(* IEC 61131-3 sources: PortalRobot/Portal_robot/Device/application/ST/ST_MULTI_TYPE, 4 files *)

(* ---- ST_MULTI_TYPE_COMMAND.st ---- *)
TYPE ST_MULTI_TYPE_COMMAND :
STRUCT
	{attribute 'symbol' := 'read'}
	xSetTypeCount         : BOOL; // Импульс изменения количества типов
	uiRequestedTypeCount : UINT; // Требуемое количество типов, 1..3
	{attribute 'symbol' := 'read'}
	xSetMachineType       : BOOL; // Импульс назначения типа станку
	uiRequestedMachine   : UINT; // Номер редактируемого станка, 1..3
	uiRequestedMachineType : UINT; // Тип, назначаемый станку
	{attribute 'symbol' := 'read'}
	xSetSlotType          : BOOL; // Импульс назначения типа слоту
	uiRequestedSlot      : UINT; // Номер редактируемого слота
	uiRequestedSlotType  : UINT; // Тип, назначаемый слоту
	{attribute 'symbol' := 'read'}
	xAutoDistribute      : BOOL; // Импульс распределения слотов пропорционально станкам
END_STRUCT
END_TYPE

(* ---- ST_MULTI_TYPE_CONFIG.st ---- *)
TYPE ST_MULTI_TYPE_CONFIG :
STRUCT
	uiTypeCount    : UINT; // Количество типов обрабатываемых деталей, 1..3
	auiMachineType : ARRAY [1..3] OF UINT; // Тип, закреплённый за каждым станком
	auiSlotType    : ARRAY [1..GVL_CELL_SETTINGS.NumberDetail] OF UINT; // Тип заготовки каждого слота
END_STRUCT
END_TYPE

(* ---- ST_MULTI_TYPE_CONFIG_STATUS.st ---- *)
TYPE ST_MULTI_TYPE_CONFIG_STATUS :
STRUCT
	xMagazineConfigAllowed   : BOOL; // Типы и распределение слотов можно менять
	xTypeCountAllowed        : BOOL; // Количество типов можно менять с применением шаблона
	axMachineTypeAllowed     : ARRAY [1..3] OF BOOL; // Назначение типа конкретному станку разрешено
	xConfigurationValid      : BOOL; // Конфигурация пригодна для автоматического цикла
	uiActiveSlotCount        : UINT; // Число слотов активной матрицы
	stWarning                : ST_WARNING_EVENT; // Последняя отклонённая команда конфигурации
END_STRUCT
END_TYPE

(* ---- ST_MULTI_TYPE_HMI.st ---- *)
TYPE ST_MULTI_TYPE_HMI :
STRUCT
	Command      : ST_MULTI_TYPE_COMMAND; // Команды конфигурации от HMI
	Config       : ST_MULTI_TYPE_CONFIG; // Фактически принятая конфигурация
	ConfigStatus : ST_MULTI_TYPE_CONFIG_STATUS; // Разрешения и диагностика конфигурации
	CycleStatus  : ST_CELL_CYCLE_STATUS; // Диагностика универсального цикла
END_STRUCT
END_TYPE
